(* IEC 61131-3 sources: plc-vscode/tests/st/test-ready/rusty/tests/lit/single/var_temp, 3 files *)

(* ---- var_temp_in_function_blocks_before_input_must_compile.st ---- *)
// RUN: (%COMPILE %s && %RUN) | %CHECK %s
FUNCTION_BLOCK Foo
    VAR_TEMP
        tmp : INT;
    END_VAR

    VAR_INPUT
        x : INT;
    END_VAR

    x := x + 1;
END_FUNCTION_BLOCK

FUNCTION main : DINT
    VAR
        fb : Foo;
    END_VAR

    fb(5);

    // CHECK: 6
    printf('%d$N', fb.x);
END_FUNCTION

(* ---- var_temp_in_function_blocks_must_compile.st ---- *)
// RUN: (%COMPILE %s && %RUN) | %CHECK %s
FUNCTION_BLOCK baseControl
    VAR_INPUT
        a_in : INT;
    END_VAR

    VAR_IN_OUT
        inoutVar : BOOL;
    END_VAR

    VAR_TEMP
        tempo : INT;
    END_VAR

    VAR_OUTPUT
        a_out :INT;
    END_VAR

    VAR

    END_VAR

    a_out := a_in + 1;

END_FUNCTION_BLOCK

FUNCTION main
   VAR
       fb : baseControl;
       fb2 : baseControl;
       dipin : BOOL;
       outVar : INT;
   END_VAR

   fb(a_in := 9, a_out => outVar, inoutVar := dipin);

   // CHECK: 10
   printf('%d$N', outVar);

   fb2(12, dipin, outVar);

   // CHECK: 13
   printf('%d$N', outVar);
END_FUNCTION

(* ---- var_temp_in_function_blocks_must_compile_when_output_has_direct_access.st ---- *)
// RUN: (%COMPILE %s && %RUN) | %CHECK %s
FUNCTION_BLOCK Foo
    VAR_TEMP
        tmp : INT;
    END_VAR

    VAR_OUTPUT
        q : BOOL;
    END_VAR

    q := TRUE;
END_FUNCTION_BLOCK

FUNCTION main : DINT
    VAR
        fb : Foo;
        result : BYTE;
    END_VAR

    fb(q => result.0);

    // CHECK: 1
    printf('%d$N', result.0);
END_FUNCTION
